// Tests for FB_HomeHold, the no-new-homing-request after a stop in the calibration sweep (#113).
FUNCTION_BLOCK FB_HomeHold_Tests EXTENDS TcUnit.FB_TestSuite
VAR
END_VAR

No_Hold_Without_Stop();
Stop_While_Homing_Holds();
Hold_Stays_After_Stop_Done();
Stop_While_Not_Homing_Does_Not_Hold();
Stop_While_Calibrated_Does_Not_Hold();
Disable_Releases_The_Hold();
Reset_Releases_The_Hold();
New_PowerOn_Releases_The_Hold();
Release_Ignored_While_Stop_Active();
Release_Without_Hold_Changes_Nothing();
StopSweep_Holds_An_Uncalibrated_Axis_Before_The_Sweep_Starts();
StopSweep_Ignored_On_A_Calibrated_Axis();
StopSweep_Wins_Over_Release_In_The_Same_Scan();
StopSweep_Hold_Ends_With_Disable();
StopSweep_Hold_Ends_With_Release_In_A_Later_Scan();

METHOD PRIVATE No_Hold_Without_Stop
VAR
	fbHold	: FB_HomeHold;
END_VAR
TEST('No_Hold_Without_Stop');
fbHold(bEnable := TRUE, bCalibrated := FALSE, bHoming := TRUE, bStopAxis := FALSE, bReset := FALSE);
AssertEquals_BOOL(Expected := FALSE, Actual := fbHold.bHold, Message := 'homing runs');
TEST_FINISHED();
END_METHOD

METHOD PRIVATE Stop_While_Homing_Holds
VAR
	fbHold	: FB_HomeHold;
END_VAR
TEST('Stop_While_Homing_Holds');
fbHold(bEnable := TRUE, bCalibrated := FALSE, bHoming := TRUE, bStopAxis := FALSE, bReset := FALSE);
fbHold(bEnable := TRUE, bCalibrated := FALSE, bHoming := TRUE, bStopAxis := TRUE, bReset := FALSE);
AssertEquals_BOOL(Expected := TRUE, Actual := fbHold.bHold, Message := 'held after the stop');
TEST_FINISHED();
END_METHOD

METHOD PRIVATE Hold_Stays_After_Stop_Done
VAR
	fbHold	: FB_HomeHold;
END_VAR
TEST('Hold_Stays_After_Stop_Done');
// bStopAxis falls on StopDone, bHomeAxis is cleared by the hold: the hold must stay while the axis is enabled
fbHold(bEnable := TRUE, bCalibrated := FALSE, bHoming := TRUE, bStopAxis := FALSE, bReset := FALSE);
fbHold(bEnable := TRUE, bCalibrated := FALSE, bHoming := TRUE, bStopAxis := TRUE, bReset := FALSE);
fbHold(bEnable := TRUE, bCalibrated := FALSE, bHoming := FALSE, bStopAxis := FALSE, bReset := FALSE);
fbHold(bEnable := TRUE, bCalibrated := FALSE, bHoming := FALSE, bStopAxis := FALSE, bReset := FALSE);
AssertEquals_BOOL(Expected := TRUE, Actual := fbHold.bHold, Message := 'still held');
TEST_FINISHED();
END_METHOD

METHOD PRIVATE Stop_While_Not_Homing_Does_Not_Hold
VAR
	fbHold	: FB_HomeHold;
END_VAR
TEST('Stop_While_Not_Homing_Does_Not_Hold');
fbHold(bEnable := TRUE, bCalibrated := FALSE, bHoming := FALSE, bStopAxis := TRUE, bReset := FALSE);
AssertEquals_BOOL(Expected := FALSE, Actual := fbHold.bHold, Message := 'no sweep, no hold');
TEST_FINISHED();
END_METHOD

METHOD PRIVATE Stop_While_Calibrated_Does_Not_Hold
VAR
	fbHold	: FB_HomeHold;
END_VAR
TEST('Stop_While_Calibrated_Does_Not_Hold');
fbHold(bEnable := TRUE, bCalibrated := TRUE, bHoming := TRUE, bStopAxis := TRUE, bReset := FALSE);
AssertEquals_BOOL(Expected := FALSE, Actual := fbHold.bHold, Message := 'calibrated');
TEST_FINISHED();
END_METHOD

METHOD PRIVATE Disable_Releases_The_Hold
VAR
	fbHold	: FB_HomeHold;
END_VAR
TEST('Disable_Releases_The_Hold');
fbHold(bEnable := TRUE, bCalibrated := FALSE, bHoming := TRUE, bStopAxis := FALSE, bReset := FALSE);
fbHold(bEnable := TRUE, bCalibrated := FALSE, bHoming := TRUE, bStopAxis := TRUE, bReset := FALSE);
fbHold(bEnable := FALSE, bCalibrated := FALSE, bHoming := FALSE, bStopAxis := FALSE, bReset := FALSE);
AssertEquals_BOOL(Expected := FALSE, Actual := fbHold.bHold, Message := 'released');
fbHold(bEnable := TRUE, bCalibrated := FALSE, bHoming := TRUE, bStopAxis := FALSE, bReset := FALSE);
AssertEquals_BOOL(Expected := FALSE, Actual := fbHold.bHold, Message := 'homing again');
TEST_FINISHED();
END_METHOD

METHOD PRIVATE Reset_Releases_The_Hold
VAR
	fbHold	: FB_HomeHold;
END_VAR
TEST('Reset_Releases_The_Hold');
fbHold(bEnable := TRUE, bCalibrated := FALSE, bHoming := TRUE, bStopAxis := FALSE, bReset := FALSE);
fbHold(bEnable := TRUE, bCalibrated := FALSE, bHoming := TRUE, bStopAxis := TRUE, bReset := FALSE);
fbHold(bEnable := TRUE, bCalibrated := FALSE, bHoming := FALSE, bStopAxis := FALSE, bReset := TRUE);
AssertEquals_BOOL(Expected := FALSE, Actual := fbHold.bHold, Message := 'released by reset');
TEST_FINISHED();
END_METHOD

METHOD PRIVATE New_PowerOn_Releases_The_Hold
VAR
	fbHold	: FB_HomeHold;
END_VAR
TEST('New_PowerOn_Releases_The_Hold');
// an automatic stop at stage 40: held, axis still enabled, reset=1 gives no bReset (#159)
fbHold(bEnable := TRUE, bCalibrated := FALSE, bHoming := TRUE, bStopAxis := FALSE, bReset := FALSE);
fbHold(bEnable := TRUE, bCalibrated := FALSE, bHoming := TRUE, bStopAxis := TRUE, bReset := FALSE);
fbHold(bEnable := TRUE, bCalibrated := FALSE, bHoming := FALSE, bStopAxis := FALSE, bReset := FALSE);
AssertEquals_BOOL(Expected := TRUE, Actual := fbHold.bHold, Message := 'held');
fbHold(bEnable := TRUE, bCalibrated := FALSE, bHoming := FALSE, bStopAxis := FALSE, bReset := FALSE, bRelease := TRUE);
AssertEquals_BOOL(Expected := FALSE, Actual := fbHold.bHold, Message := 'released by the new power-on');
TEST_FINISHED();
END_METHOD

METHOD PRIVATE Release_Ignored_While_Stop_Active
VAR
	fbHold	: FB_HomeHold;
END_VAR
TEST('Release_Ignored_While_Stop_Active');
fbHold(bEnable := TRUE, bCalibrated := FALSE, bHoming := TRUE, bStopAxis := FALSE, bReset := FALSE);
fbHold(bEnable := TRUE, bCalibrated := FALSE, bHoming := TRUE, bStopAxis := TRUE, bReset := FALSE, bRelease := TRUE);
AssertEquals_BOOL(Expected := TRUE, Actual := fbHold.bHold, Message := 'a running stop is not cut through');
TEST_FINISHED();
END_METHOD

METHOD PRIVATE Release_Without_Hold_Changes_Nothing
VAR
	fbHold	: FB_HomeHold;
END_VAR
TEST('Release_Without_Hold_Changes_Nothing');
fbHold(bEnable := TRUE, bCalibrated := FALSE, bHoming := TRUE, bStopAxis := FALSE, bReset := FALSE, bRelease := TRUE);
AssertEquals_BOOL(Expected := FALSE, Actual := fbHold.bHold, Message := 'no hold');
TEST_FINISHED();
END_METHOD

METHOD PRIVATE StopSweep_Holds_An_Uncalibrated_Axis_Before_The_Sweep_Starts
VAR
	fbHold	: FB_HomeHold;
END_VAR
TEST('StopSweep_Holds_An_Uncalibrated_Axis_Before_The_Sweep_Starts');
// #198: the stop arrives before bHomeAxis is set (tonReady, or the scans after a reset)
fbHold(bEnable := TRUE, bCalibrated := FALSE, bHoming := FALSE, bStopAxis := FALSE, bReset := FALSE, bStopSweep := TRUE);
AssertEquals_BOOL(Expected := TRUE, Actual := fbHold.bHold, Message := 'held');
fbHold(bEnable := TRUE, bCalibrated := FALSE, bHoming := FALSE, bStopAxis := FALSE, bReset := FALSE, bStopSweep := FALSE);
AssertEquals_BOOL(Expected := TRUE, Actual := fbHold.bHold, Message := 'still held');
TEST_FINISHED();
END_METHOD

METHOD PRIVATE StopSweep_Ignored_On_A_Calibrated_Axis
VAR
	fbHold	: FB_HomeHold;
END_VAR
TEST('StopSweep_Ignored_On_A_Calibrated_Axis');
fbHold(bEnable := TRUE, bCalibrated := TRUE, bHoming := FALSE, bStopAxis := FALSE, bReset := FALSE, bStopSweep := TRUE);
AssertEquals_BOOL(Expected := FALSE, Actual := fbHold.bHold, Message := 'calibrated axis not held');
TEST_FINISHED();
END_METHOD

METHOD PRIVATE StopSweep_Wins_Over_Release_In_The_Same_Scan
VAR
	fbHold	: FB_HomeHold;
END_VAR
TEST('StopSweep_Wins_Over_Release_In_The_Same_Scan');
fbHold(bEnable := TRUE, bCalibrated := FALSE, bHoming := FALSE, bStopAxis := FALSE, bReset := FALSE, bRelease := TRUE, bStopSweep := TRUE);
AssertEquals_BOOL(Expected := TRUE, Actual := fbHold.bHold, Message := 'held');
TEST_FINISHED();
END_METHOD

METHOD PRIVATE StopSweep_Hold_Ends_With_Disable
VAR
	fbHold	: FB_HomeHold;
END_VAR
TEST('StopSweep_Hold_Ends_With_Disable');
fbHold(bEnable := TRUE, bCalibrated := FALSE, bHoming := FALSE, bStopAxis := FALSE, bReset := FALSE, bStopSweep := TRUE);
fbHold(bEnable := FALSE, bCalibrated := FALSE, bHoming := FALSE, bStopAxis := FALSE, bReset := FALSE, bStopSweep := FALSE);
AssertEquals_BOOL(Expected := FALSE, Actual := fbHold.bHold, Message := 'released by the disable');
TEST_FINISHED();
END_METHOD

METHOD PRIVATE StopSweep_Hold_Ends_With_Release_In_A_Later_Scan
VAR
	fbHold	: FB_HomeHold;
END_VAR
TEST('StopSweep_Hold_Ends_With_Release_In_A_Later_Scan');
fbHold(bEnable := TRUE, bCalibrated := FALSE, bHoming := FALSE, bStopAxis := FALSE, bReset := FALSE, bStopSweep := TRUE);
fbHold(bEnable := TRUE, bCalibrated := FALSE, bHoming := FALSE, bStopAxis := FALSE, bReset := FALSE, bRelease := TRUE, bStopSweep := FALSE);
AssertEquals_BOOL(Expected := FALSE, Actual := fbHold.bHold, Message := 'released by a new power-on');
TEST_FINISHED();
END_METHOD

END_FUNCTION_BLOCK

(* stored: Version 1.1.0.1, ProductVersion 3.1.4024.15
   POU FB_HomeHold_Tests: Id {6bb4a0fd-8b06-4947-b443-64dcd332a1b6}, SpecialFunc None
   Method No_Hold_Without_Stop: Id {e618cb85-d147-45e8-af5c-d7c17a1c1091}
   Method Stop_While_Homing_Holds: Id {5540370c-90bd-4706-bb24-be044a49aaec}
   Method Hold_Stays_After_Stop_Done: Id {de167aeb-f4f2-4ff9-b738-fd11f0c3ce0d}
   Method Stop_While_Not_Homing_Does_Not_Hold: Id {50b1c3a5-a03d-446e-a1c8-3f2c2f006b58}
   Method Stop_While_Calibrated_Does_Not_Hold: Id {d4107741-efd3-478e-8bb1-c6be2b97eeab}
   Method Disable_Releases_The_Hold: Id {aa073480-334e-4252-8f13-7e00f11f97a3}
   Method Reset_Releases_The_Hold: Id {28edd587-aed6-409a-8338-2eccfa7208c5}
   Method New_PowerOn_Releases_The_Hold: Id {c1a7e302-5b94-4d1f-8a60-3e92b7d0f411}
   Method Release_Ignored_While_Stop_Active: Id {7e50b9d4-2a13-4c68-b0f5-91d8c3a4e627}
   Method Release_Without_Hold_Changes_Nothing: Id {e94d2f81-0c7b-4a35-9d16-b8a5e0f3c752}
   Method StopSweep_Holds_An_Uncalibrated_Axis_Before_The_Sweep_Starts: Id {c8e4d888-cf30-46f7-9257-b533bf879c95}
   Method StopSweep_Ignored_On_A_Calibrated_Axis: Id {d5cc4f73-8d57-49c4-95bc-ea4167a5039d}
   Method StopSweep_Wins_Over_Release_In_The_Same_Scan: Id {11e7a50a-4407-4d05-b7bd-7c53a2f391e4}
   Method StopSweep_Hold_Ends_With_Disable: Id {7a273dbf-c555-4785-93f3-7e97d24eab83}
   Method StopSweep_Hold_Ends_With_Release_In_A_Later_Scan: Id {5de5d511-f0ce-4959-be2c-fa3d49135d43} *)
